(*
SPDX-FileCopyrightText: © 2026 Oleksandr Tiutyk <trofimich@gmail.com>
SPDX-License-Identifier: MIT
License: https://opensource.org/license/mit
*)

(*!
<summary>Provides fluent assertions on a copied LDATE value.</summary>
<description>
Copies actual into persistent instance storage before the entry method returns; literals and expression
results therefore remain valid throughout the immediate chain. Owns no heap allocation or pointed-to resource.
The message prefixes every failure until the next preparation. Finish one chain before starting another on
the owning Assertions provider. Use only from the owning test callback on one task, without reentry.
Obtain this context from the owning provider; direct unprepared use is unsupported.
Expected arguments use the declared IEC type; ordinary compiler conversions happen before comparison.
This context does not depend on another assertion context.
Object metadata is available before preparation; inherited equality compares instance identity.
</description>
*)

{attribute 'no_explicit_call' := 'do not call this function block directly'}
FUNCTION_BLOCK LongDateAssertionContext EXTENDS TOF_Core.Object
VAR_STAT
	{attribute 'hide'}
	_ClassName : STRING := __POUNAME();
END_VAR
VAR
	_Actual : LDATE;
	_TestCase : ITestCase;
	_Message : WSTRING(255);
END_VAR

(*!
<summary>Provides the implementation class name.</summary>
<description>
Borrowed read-only reference to compiler-initialized storage, valid throughout the instance lifetime.
Do not modify the returned reference; no ownership is transferred.
</description>
*)
{attribute 'monitoring' := 'call'}
PROPERTY ClassName : REFERENCE TO STRING
GET
ClassName REF= _ClassName;
END_GET
END_PROPERTY

(*!
<summary>Asserts that the actual value is strictly greater than expected.</summary>
<description>
Records failure without interrupting the callback; preserves the message for the rest of the chain.
</description>
<param name="expected">Expected value converted by the compiler to LDATE.</param>
*)
METHOD FINAL IsGreaterThan : REFERENCE TO LongDateAssertionContext
VAR_INPUT
	expected : LDATE;
END_VAR
IF _Actual <= expected THEN
	failComparison(
		expected := expected,
		expectation := "Expected value > "
	);
END_IF

IsGreaterThan REF= THIS^;
END_METHOD

(*!
<summary>Asserts that the actual value meets the inclusive lower boundary.</summary>
<description>
Records failure without interrupting the callback; preserves the message for the rest of the chain.
</description>
<param name="expected">Expected value converted by the compiler to LDATE.</param>
*)
METHOD FINAL IsGreaterThanOrEquals : REFERENCE TO LongDateAssertionContext
VAR_INPUT
	expected : LDATE;
END_VAR
IF _Actual < expected THEN
	failComparison(
		expected := expected,
		expectation := "Expected value >= "
	);
END_IF

IsGreaterThanOrEquals REF= THIS^;
END_METHOD

(*!
<summary>Asserts that the actual value is strictly less than expected.</summary>
<description>
Records failure without interrupting the callback; preserves the message for the rest of the chain.
</description>
<param name="expected">Expected value converted by the compiler to LDATE.</param>
*)
METHOD FINAL IsLessThan : REFERENCE TO LongDateAssertionContext
VAR_INPUT
	expected : LDATE;
END_VAR
IF _Actual >= expected THEN
	failComparison(
		expected := expected,
		expectation := "Expected value < "
	);
END_IF

IsLessThan REF= THIS^;
END_METHOD

(*!
<summary>Asserts that the actual value meets the inclusive upper boundary.</summary>
<description>
Records failure without interrupting the callback; preserves the message for the rest of the chain.
</description>
<param name="expected">Expected value converted by the compiler to LDATE.</param>
*)
METHOD FINAL IsLessThanOrEquals : REFERENCE TO LongDateAssertionContext
VAR_INPUT
	expected : LDATE;
END_VAR
IF _Actual > expected THEN
	failComparison(
		expected := expected,
		expectation := "Expected value <= "
	);
END_IF

IsLessThanOrEquals REF= THIS^;
END_METHOD

(*!
<summary>Provides the library namespace.</summary>
<description>
Borrowed read-only reference to the compiler-initialized namespace, valid throughout the instance lifetime.
Do not modify the returned reference; no ownership is transferred.
</description>
*)
{attribute 'monitoring' := 'call'}
PROPERTY NamespaceName : REFERENCE TO STRING
GET
NamespaceName REF= CurrentNamespace.Name;
END_GET
END_PROPERTY

(*!
<summary>Asserts inequality with the expected value.</summary>
<description>
Records failure without interrupting the callback; preserves the message for the rest of the chain.
</description>
<param name="expected">Expected value converted by the compiler to LDATE.</param>
*)
METHOD FINAL NotToBe : REFERENCE TO LongDateAssertionContext
VAR_INPUT
	expected : LDATE;
END_VAR
IF _Actual = expected THEN
	failComparison(
		expected := expected,
		expectation := "Expected value not to be: "
	);
END_IF

NotToBe REF= THIS^;
END_METHOD

(*!
<summary>Copies the actual operand and replaces the chain-wide message.</summary>
<description>
Called by the owning Assertions provider after it verifies the running test case.
No pointer to this method's input storage is retained. The receiver is borrowed until the next preparation;
the owning provider keeps it alive throughout the immediate chain.
</description>
<param name="actual">Value copied into this context.</param>
<param name="testCase">Borrowed failure receiver for the immediate chain.</param>
<param name="message">Copied diagnostic prefix, including empty to clear the previous prefix.</param>
*)
METHOD INTERNAL FINAL Prepare
VAR_INPUT
	actual : LDATE;
	testCase : ITestCase;
	message : WSTRING(255);
END_VAR
_Actual := actual;
_TestCase := testCase;
_Message := message;
END_METHOD

(*!
<summary>Reports the byte size of this concrete instance.</summary>
<description>
Includes inline fields and nested instances, but excludes separately allocated payloads.
Obtaining the size does not transfer ownership or validate an arbitrary address.
</description>
*)
{attribute 'monitoring' := 'call'}
PROPERTY SelfSize : ULINT
GET
SelfSize := XSIZEOF(THIS^);
END_GET
END_PROPERTY

(*!
<summary>Asserts equality with the expected value.</summary>
<description>
Records failure without interrupting the callback; preserves the message for the rest of the chain.
</description>
<param name="expected">Expected value converted by the compiler to LDATE.</param>
*)
METHOD FINAL ToBe : REFERENCE TO LongDateAssertionContext
VAR_INPUT
	expected : LDATE;
END_VAR
IF _Actual <> expected THEN
	failComparison(
		expected := expected,
		expectation := "Expected: "
	);
END_IF

ToBe REF= THIS^;
END_METHOD

(*!
<summary>Formats a failed typed predicate and reports it with the chain message.</summary>
<description>
Does not change operands or chain state. The receiver retains its first failure. Reporting exceptions
propagate to the enclosing test callback handler; an unprepared receiver is a configuration error.
</description>
<param name="expected">Typed expected operand used only for this diagnostic.</param>
<param name="expectation">Prefix identifying the failed predicate.</param>
*)
METHOD PRIVATE failComparison
VAR_INPUT
	expected : LDATE;
	expectation : WSTRING(40);
END_VAR
VAR
	actualText : WSTRING(255);
	expectedText : WSTRING(255);
	diagnostic : TOF_Core.ERROR_MESSAGE;
END_VAR
actualText := TO_WSTRING(_Actual);
expectedText := TO_WSTRING(expected);

diagnostic := TOF_Core.WideStrings.Concat255(
	expectation,
	expectedText,
	", but was: ",
	actualText
);

TestServices.ReportAssertionFailure(
	testCase := _TestCase,
	message := _Message,
	sourceClassName := ClassName,
	defaultMessage := diagnostic
);
END_METHOD

END_FUNCTION_BLOCK

(* stored: Version 1.1.0.1
   POU LongDateAssertionContext: Id {e52335c9-ec4b-43fe-8d63-12f6ce621b6a}, SpecialFunc None
   Folder Service methods: Id {1544f12f-2f21-41bf-bede-105db13f5bfd}
   Property ClassName: Id {9fd2e6fa-5009-48f5-a8b3-f0fb37a26d4e}
   Get Get: Id {7319c41e-05fc-410e-9fa1-567cf9b1f494}
   Method IsGreaterThan: Id {ea6d2d10-dcd4-4e73-9040-12e2eef3f506}
   Method IsGreaterThanOrEquals: Id {b3022f54-7d95-42a7-932f-59d1ba691138}
   Method IsLessThan: Id {03eef457-a0a1-4a59-9621-3649bf63061f}
   Method IsLessThanOrEquals: Id {9f5f7e33-3818-46d7-acbc-3c5a52a18c06}
   Property NamespaceName: Id {2c728f37-e2df-4ae9-8124-2c9bbfb1b120}
   Get Get: Id {c03cef7e-7e40-4f84-a15b-1d7f531202db}
   Method NotToBe: Id {910c30d2-5b16-4160-8d27-c4d993bfe851}
   Method Prepare: Id {638e39d9-c400-45f7-ba62-c455b5434aa8}
   Property SelfSize: Id {f32afeaf-1c70-489b-afcd-3044622da94d}
   Get Get: Id {c06ce974-d674-4478-8045-860171041966}
   Method ToBe: Id {f55c8ffd-5f43-4a66-908f-c9a57ba86921}
   Method failComparison: Id {15223af9-a9d9-416a-9199-8c41b6022287} *)
